FUNCTION_BLOCK IO_RouteAI (* Picks the way an IO block reaches its signal from the Address (a Pi line, a local IO handle, Modbus or simulated) and passes values through that way only. Technical: Backend router for IO_AI; Address: 'gpio[chip:line(:pull_up|:pull_down)(:active_low)]' or 'pwm[chip:channel:period_ns]' a Raspberry Pi's line, set up here; 'modbus[...]' a Modbus CLIENT ID; 'sim' simulated; another name a local IO handle set up elsewhere (IX/QX PARAMS); empty: not connected (QO = FALSE) *)
  (* Standard: 61499-2 *)
  (* Version 0.1, 2026-09-28, Project contributors, AAU Smart Production Lab *)
  PACKAGE modlib;
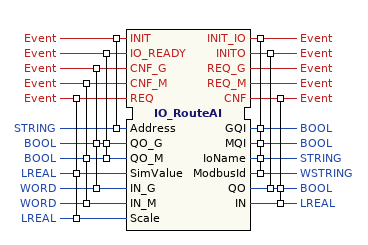
  EVENT_INPUT
    INIT WITH Address; (* Work out from Address how the point is reached *)
    IO_READY WITH QO_G, QO_M; (* The line, the local IO block and the Modbus client are initialised *)
    CNF_G WITH QO_G, IN_G; (* The local IO block answered *)
    CNF_M WITH QO_M, IN_M; (* The Modbus client answered *)
    REQ WITH SimValue, Scale; (* Access the point *)
  END_EVENT
  EVENT_OUTPUT
    INIT_IO WITH GQI, MQI, IoName, ModbusId; (* Set up the line, the local IO block and the Modbus client (each only if it is the way) *)
    INITO WITH QO; (* Initialised: QO says whether the point is reachable *)
    REQ_G; (* Access the point through the local IO block (IX/QX/IW/QW) *)
    REQ_M; (* Access the point through the Modbus client *)
    CNF WITH QO, IN; (* Done: QO says whether it worked *)
  END_EVENT
  VAR_INPUT
    Address : STRING; (* Where the point is: 'gpio[chip:line(:pull_up|:pull_down)(:active_low)]', 'pwm[chip:channel:period_ns]', 'modbus[...]', 'sim', or an IO handle's name; empty: not connected *)
    QO_G : BOOL; (* The local IO block works *)
    QO_M : BOOL; (* The Modbus client works *)
    SimValue : LREAL; (* The value read when the address is 'sim' *)
    IN_G : WORD; (* The raw value read through the local IO block *)
    IN_M : WORD; (* The raw value read through Modbus *)
    Scale : LREAL := 1.0; (* Engineering value per raw count *)
  END_VAR
  VAR_OUTPUT
    GQI : BOOL; (* Use the local IO block *)
    MQI : BOOL; (* Use the Modbus client *)
    IoName : STRING; (* The local IO handle's name (PARAMS of IX/QX/IW/QW) *)
    ModbusId : WSTRING; (* The Modbus CLIENT's ID *)
    QO : BOOL; (* The point is reachable, the last access worked *)
    IN : LREAL; (* The value read (an analog one scaled) *)
  END_VAR
  VAR
    Backend : USINT;
  END_VAR
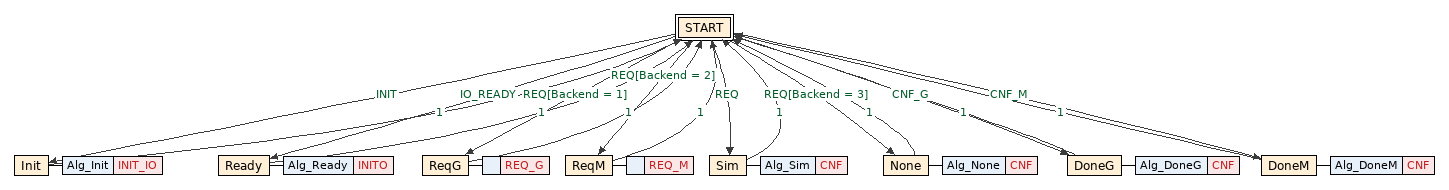
  EC_STATES
    START;
    Init : Alg_Init -> INIT_IO;
    Ready : Alg_Ready -> INITO;
    ReqG : -> REQ_G;
    ReqM : -> REQ_M;
    Sim : Alg_Sim -> CNF;
    None : Alg_None -> CNF;
    DoneG : Alg_DoneG -> CNF;
    DoneM : Alg_DoneM -> CNF;
  END_STATES
  EC_TRANSITIONS
    START TO Init := INIT;
    Init TO START := 1;
    START TO Ready := IO_READY;
    Ready TO START := 1;
    START TO ReqG := REQ[Backend = 1];
    START TO ReqM := REQ[Backend = 2];
    START TO None := REQ[Backend = 3];
    START TO Sim := REQ;
    START TO DoneG := CNF_G;
    START TO DoneM := CNF_M;
    ReqG TO START := 1;
    ReqM TO START := 1;
    Sim TO START := 1;
    None TO START := 1;
    DoneG TO START := 1;
    DoneM TO START := 1;
  END_TRANSITIONS
  ALGORITHM Alg_Init IN ST:
Backend := 3;
IF Address = 'sim' THEN
  Backend := 0;
ELSIF LEFT(Address, 7) = 'modbus[' THEN
  Backend := 2;
  ModbusId := STRING_TO_WSTRING(Address);
ELSIF LEN(Address) > 0 THEN
  Backend := 1;
  IoName := Address;
END_IF;
GQI := Backend = 1;
MQI := Backend = 2;
  END_ALGORITHM
  ALGORITHM Alg_Ready IN ST:
QO := (Backend = 0) OR ((Backend = 1) AND QO_G) OR ((Backend = 2) AND QO_M);
  END_ALGORITHM
  ALGORITHM Alg_Sim IN ST:
QO := TRUE;
IN := SimValue;
  END_ALGORITHM
  ALGORITHM Alg_None IN ST:
QO := FALSE;
  END_ALGORITHM
  ALGORITHM Alg_DoneG IN ST:
QO := QO_G;
IN := UINT_TO_LREAL(WORD_TO_UINT(IN_G)) * Scale;
  END_ALGORITHM
  ALGORITHM Alg_DoneM IN ST:
QO := QO_M;
IN := UINT_TO_LREAL(WORD_TO_UINT(IN_M)) * Scale;
  END_ALGORITHM
END_FUNCTION_BLOCK
